TYPE ST_SrmKinematics :
STRUCT
    lrVeloX  : LREAL;   // travel
    lrAccelX : LREAL;
    lrVeloY  : LREAL;   // hoist
    lrAccelY : LREAL;
    lrVeloZ  : LREAL;   // telescopic fork
    lrAccelZ : LREAL;
END_STRUCT
END_TYPE

(* stored: Version 1.1.0.1
   DUT ST_SrmKinematics: Id {82b22a17-5091-40dc-8654-72c5bc060c9e} *)
